Fanuc KAREL source: KX00006.KL

PROGRAM KX00006
%NOLOCKGROUP
VAR
  I: INTEGER
  J: INTEGER
  B: BOOLEAN
  F: FILE
  S: STRING[80]
  P: XYZWPR
BEGIN
  PULSE DOUT[1] FOR 100
END KX00006
